TYPE "st_Station_Hp_Instruments"
VERSION : 0.1
   STRUCT
      Zone2_FM1 { ExternalAccessible := 'False'; ExternalVisible := 'False'; ExternalWritable := 'False'; S7_SetPoint := 'False'} : "st_Station_Hp_InstrumentPosition";
      Zone2_FM2 { ExternalAccessible := 'False'; ExternalVisible := 'False'; ExternalWritable := 'False'; S7_SetPoint := 'False'} : "st_Station_Hp_InstrumentPosition";
      Zone2_FM3 { ExternalAccessible := 'False'; ExternalVisible := 'False'; ExternalWritable := 'False'; S7_SetPoint := 'False'} : "st_Station_Hp_InstrumentPosition";
      Zone2_FM4 { ExternalAccessible := 'False'; ExternalVisible := 'False'; ExternalWritable := 'False'; S7_SetPoint := 'False'} : "st_Station_Hp_InstrumentPosition";
      Zone3_FM1 { ExternalAccessible := 'False'; ExternalVisible := 'False'; ExternalWritable := 'False'; S7_SetPoint := 'False'} : "st_Station_Hp_InstrumentPosition";
      Zone3_FM2 { ExternalAccessible := 'False'; ExternalVisible := 'False'; ExternalWritable := 'False'; S7_SetPoint := 'False'} : "st_Station_Hp_InstrumentPosition";
      Zone3_FM3 { ExternalAccessible := 'False'; ExternalVisible := 'False'; ExternalWritable := 'False'; S7_SetPoint := 'False'} : "st_Station_Hp_InstrumentPosition";
      Zone3_FM4 { ExternalAccessible := 'False'; ExternalVisible := 'False'; ExternalWritable := 'False'; S7_SetPoint := 'False'} : "st_Station_Hp_InstrumentPosition";
      Zone1_Pt1 { ExternalAccessible := 'False'; ExternalVisible := 'False'; ExternalWritable := 'False'; S7_SetPoint := 'False'} : "st_Station_Hp_InstrumentPosition";
      Zone2_Pt1 { ExternalAccessible := 'False'; ExternalVisible := 'False'; ExternalWritable := 'False'; S7_SetPoint := 'False'} : "st_Station_Hp_InstrumentPosition";
      Zone2_Pt2 { ExternalAccessible := 'False'; ExternalVisible := 'False'; ExternalWritable := 'False'; S7_SetPoint := 'False'} : "st_Station_Hp_InstrumentPosition";
      Zone3_Pt1 { ExternalAccessible := 'False'; ExternalVisible := 'False'; ExternalWritable := 'False'; S7_SetPoint := 'False'} : "st_Station_Hp_InstrumentPosition";
      Zone3_Pt2 { ExternalAccessible := 'False'; ExternalVisible := 'False'; ExternalWritable := 'False'; S7_SetPoint := 'False'} : "st_Station_Hp_InstrumentPosition";
      Zone1_Vacuummeter1 { ExternalAccessible := 'False'; ExternalVisible := 'False'; ExternalWritable := 'False'; S7_SetPoint := 'False'} : "st_Station_Hp_InstrumentPosition";
      Zone2_Vacuummeter1 { ExternalAccessible := 'False'; ExternalVisible := 'False'; ExternalWritable := 'False'; S7_SetPoint := 'False'} : "st_Station_Hp_InstrumentPosition";
      Zone2_Vacuummeter2 { ExternalAccessible := 'False'; ExternalVisible := 'False'; ExternalWritable := 'False'; S7_SetPoint := 'False'} : "st_Station_Hp_InstrumentPosition";
      Zone3_Vacuummeter1 { ExternalAccessible := 'False'; ExternalVisible := 'False'; ExternalWritable := 'False'; S7_SetPoint := 'False'} : "st_Station_Hp_InstrumentPosition";
      Zone3_Vacuummeter2 { ExternalAccessible := 'False'; ExternalVisible := 'False'; ExternalWritable := 'False'; S7_SetPoint := 'False'} : "st_Station_Hp_InstrumentPosition";
      Zone1_FM1 { ExternalAccessible := 'False'; ExternalVisible := 'False'; ExternalWritable := 'False'; S7_SetPoint := 'False'} : "st_Station_Hp_InstrumentPosition";
      Zone1_FM2 { ExternalAccessible := 'False'; ExternalVisible := 'False'; ExternalWritable := 'False'; S7_SetPoint := 'False'} : "st_Station_Hp_InstrumentPosition";
   END_STRUCT;

END_TYPE

